(* IEC 61131-3 sources: NachHouse_TST/ROOM_API_PILOT/CODEX_BACKUP_20260826_2304, 1 file *)

(* ---- prgMain.ST ---- *)
PROGRAM prgMain
  VAR_INPUT
  END_VAR
  VAR_OUTPUT
  END_VAR
  VAR
  END_VAR
  VAR_TEMP
  END_VAR

END_PROGRAM
